// System API/SYS/API/bds_sys_do
///This function set the digital system output to the given state.
///
///=======
/// Remarks:
///=======
///    + The function is just used for the reactivation of the shunt after the elapsed recovery time and therefore a switch off is not necessary. 
///    + The |GVL_sys| is given for usage of defines.
///    + Import the bds_rts_ec.xml to use the enums. (Refer example below).
///
///----------
/// FFI:
///----------
///This API can be used in trusted partitions only. See Freedom from Interference (FFI) concept for more details.
///
///==================================================================		  			===================================================================================================
///Return value    								  									Description
///==================================================================		  			===================================================================================================
///16#00																				No error.
///16#01																				A parameter is invalid.
///16#02																				Function call was erroneous.
///16#03																				Shunt activation is not enabled.
///16#04																				Recovery time is not elapsed.
///
///==================================================================		   			===================================================================================================
///
///=======
///Code Example:
///=======
///============================================================================
///
///PROGRAM PLC_PRG
///
///VAR
///
///	status_u8: UISNT := 16#00; 
/// 
///	Init_flag_u8:USINT:=0;
///
///END_VAR
///
///  
///IF(Init_flag_u8=0) THEN (*To make api call once in application*)
///
///	(* reactivate the shunt after detection of a short circuit to battery *)
///	
///	status_u8 := bds_sys_do(bds_sys_do_signal_te.SHUNT1_EN, STD_ACTIVE);
///	
///	Init_flag_u8:=1;
///  
///END_IF
///
///============================================================================
{attribute 'external_name' := 'cmp_rts_bds_sys_do'}
FUNCTION bds_sys_do : USINT
VAR_INPUT
	///The assigned signal name.
	signal_e: UINT;
	///States of the sensor supply.
	///
	///    + STD_OFF - Disable the digital output,
	///    + STD_ON   - Enable the digital output.
	state_u8: USINT;
END_VAR

END_FUNCTION

// I/O API/IN legacy/API/bds_in_aid
///Get the analog voltage of the input as state.
///
///=======
/// Remarks:
///=======
///    + The evaluation of the state (and also the diagnosis OR (out of range)) is only possible with the configuration of the state thresholds. ( see |bds_in_aid_cfg|).
///
///----------
/// FFI:
///----------
///This API can be used in trusted partitions only. See Freedom from Interference (FFI) concept for more details.
///
///	
///==================================================================		  			===================================================================================================
///Return value    								  									Description
///==================================================================		  			===================================================================================================
///0																					No error
///1																					Invalid parameter
///2																					Function call was erroneous
///3																					Thresholds are not configured
///
///==================================================================		   			===================================================================================================
///
///=======
///Code Example:
///=======
///============================================================================
///
///PROGRAM appl_10ms_task
///  VAR
///  
///    stK59_u8: USINT := 16#00;
///  END_VAR
///
///  (* get the state of input K59 *)
///  
///  bds_in_aid(bds_in_aiv_signal_te.K59, ADR(stK59_u8));
///END
///
///============================================================================
{attribute 'external_name' := 'cmp_rts_bds_in_aid'}
FUNCTION bds_in_aid : USINT
VAR_INPUT
	///The signal name that is assigned to the respective pin configured as voltage input
	signal_e: UINT;
	///Storage address of the state.
	///	
	///States:
	///    + 0 : OFF
	///    + 1 : ON
	state_pu8: POINTER TO USINT;
END_VAR

END_FUNCTION

// I/O API/IN legacy/API/bds_in_aid_cfg
///Configure the state thresholds voltages of the input.
///
///=======
/// Remarks:
///=======
///    + The evaluation of the state and also the diagnosis of out of range (OR) is only possible with the configuration of the state thresholds (see also Configure a digital input.)
///	    + With a diagnosis threshold range of 150 to 4850mV or 150 to 19850mV or 150 to 39850mV, the corresponding state threshold range for the configurable inputs are defined from 300 to 4700mV or 300 to 19700mV or 300 to 39700mV depending upon the configuration.
///	    + With a diagnosis threshold range of 150 to 29850mV the state threshold range for the fixed inputs is defined from 300 to 29700mV. 
///    + For more information see |bds_in_aiv_getStatus|. 
///    + The AID_cfg  function is not recommended for the discrete inputs that have pull-up to battery (14K7) and pull-down (80K). 
///    + For discrete inputs, the thresholds depend on the battery voltage. It is recommended to do the evaluation of the states in ASW by reading the current battery voltage for a particular input and to calculate the appropriate thresholds for that battery voltage.
///
///----------
/// FFI:
///----------
///This API can be used in trusted partitions only. See Freedom from Interference (FFI) concept for more details.
///
///	
///==================================================================		  			===================================================================================================
///Return value    								  									Description
///==================================================================		  			===================================================================================================
///0																					No error
///1																					Invalid parameter
///
///==================================================================		   			===================================================================================================
///
///=======
///Code Example:
///=======
///============================================================================
///
///PROGRAM appl_10ms_task
///  VAR
///  
///  END_VAR
///
/// (* configure the state thresholds of input K59 *)
///
///  bds_in_aid_cfg(bds_in_aiv_signal_te.K59, 3000, 2000);
///END
///
///============================================================================
{attribute 'external_name' := 'cmp_rts_bds_in_aid_cfg'}
FUNCTION bds_in_aid_cfg : USINT
VAR_INPUT
	///The signal name that is assigned to the respective pin configured as voltage input
	signal_e: UINT;
	///Upper state threshold [mV].
	///
	///Range:
	///
	///Configurable inputs:
	///300 to 4700 / 300 to 19700 /300 to 39700
	///
	///Fixed inputs:
	///300 to 29700 
	///
	///Note:
	///upperThreshold_u16 > lowerThreshold_u16
	upperThreshold_u16: UINT;
	///Lower diagnosis threshold [mV].
	///
	///Range:
	///
	///Configurable inputs:
	///300 to 4700 / 300 to 19700 / 300 to 39700
	///
	///Fixed inputs:
	///300 to 29700
	///
	///Note:
	///lowerThreshold_u16 < upperThreshold_u16
	lowerThreshold_u16: UINT;
END_VAR

END_FUNCTION

// I/O API/IN legacy/API/bds_in_aiv
///Provides the analog voltage of the input.
///
///=======
/// Remarks:
///=======
///The voltage range of the inputs depends on the input type and the input configuration using eC (easyConfig). (see also |bds_in_aiv_cfg| and |bds_in_aid_cfg|).
///	   + Based on the configuration, the measurement range of the input  can  be  0 to 5000mV or 0 to 20000mV or 0 to 40000mV 
///	   + The measurement range of the routed input via the input device is 0 to 5000mV, see also Analog voltage aquisition.
///	   + The measurement range of the discrete inputs is 0 to 33000mV or 0 to 5000 mV
///
///
///----------
/// FFI:
///----------
///This API can be used in trusted partitions only. See Freedom from Interference (FFI) concept for more details.
///
///==================================================================		  			===================================================================================================
///Return value    								  									Description
///==================================================================		  			===================================================================================================
///0																					No error
///1																					Invalid parameter
///
///==================================================================		   			===================================================================================================
///
///
///=======
///Code Example:
///=======
///============================================================================
///
///PROGRAM appl_10ms_task
///  VAR
///  
///    mV_K59_u16: UINT := 16#00;
///  END_VAR
///
/// (* get the voltage of input K59 *)
///
///  bds_in_aiv(bds_in_aiv_signal_te.K59, ADR(mV_K59_u16));
///END
///
///============================================================================
{attribute 'external_name' := 'cmp_rts_bds_in_aiv'}
FUNCTION bds_in_aiv : USINT
VAR_INPUT
	///The signal name that is assigned to the respective pin configured as voltage input
	signal_e: UINT;
	///Storage address of the value.
	///
	///Range:
	///0 to 40000  [mV]
	value_pu16: POINTER TO UINT;
END_VAR

END_FUNCTION

// I/O API/IN legacy/API/bds_in_aiv_cfg
///Configures the diagnosis thresholds voltages of the input.
///
///=======
/// Remarks:
///=======
///   + The diagnosis is only possible after the configuration of the diagnosis thresholds. 
///	   + Depending on the configuration, the diagnosis threshold range for the configurable inputs can be from 150 to 4850 or 150 to 19850 or 150 to 39850mV.
///	   + The diagnosis threshold range for the fixed inputs ranges is from 150 to 29850mV or 150 to 4850 mV.
///   + For more information see |bds_in_aiv_getStatus|.
///   + This function should be called only once in the application.
///	
///
///----------
/// FFI:
///----------
///This API can be used in trusted partitions only. See Freedom from Interference (FFI) concept for more details.
///
///==================================================================		  			===================================================================================================
///Return value    								  									Description
///==================================================================		  			===================================================================================================
///0																					No error
///1																					Invalid parameter
///2																					Function call was erroneous.
///
///==================================================================		   			===================================================================================================
///
///=======
///Code Example:
///=======
///============================================================================
///
///PROGRAM PLC_PRG
///
///  VAR
///  
///	Init_flag_u8:USINT:=0;
/// 
///  END_VAR
///
///IF(Init_flag_u8=0) THEN (*To make api call once in application*)
///
///	(* configure diagnosis thresholds of input K59 *)
///	
///	bds_in_aiv_cfg(bds_in_aiv_signal_te.K59, 4850, 150);
///	
///	Init_flag_u8:=1;
///  
///END_IF
///
///============================================================================
{attribute 'external_name' := 'cmp_rts_bds_in_aiv_cfg'}
FUNCTION bds_in_aiv_cfg : USINT
VAR_INPUT
	///The signal name that is assigned to the respective pin configured as voltage input.
	signal_e: UINT;
	///Higher diagnosis threshold in [mV].
	///
	///Range:
	///
	///Configurable inputs:
	///150 to 4850 / 150 to 19850 / 150 to 39850
	///
	///Fixed inputs:
	///150 to 29850
	///
	///Note:
	///upperThreshold_u16 > lowerThreshold_u16
	upperThreshold_u16: UINT;
	///Lower diagnosis threshold in [mV].
	///
	///Range:
	///
	///Configurable inputs:
	///150 to 4850 / 150 to 19850 / 150 to 39850
	///
	///Fixed inputs:
	///150 to 29850
	///
	///Note:
	///lowerThreshold_u16 < upperThreshold_u16
	lowerThreshold_u16: UINT;
END_VAR

END_FUNCTION

// I/O API/IN legacy/API/bds_in_phase
///Provides the signal and the phase information of a channel (consist of a primary and a secondary frequency signal).
///
///=======
/// Remarks:
///=======
///   + The phase measurement for a phase channel can be configured through easyConfig and is automatically enabled during the start up of the ECU.
///   + All frequency inputs can be grouped to predefined input pairs.
///   + For information about the signal acquisition see Frequency aquisition.
///   + Following signal information is available: 
///	   + Frequency information of the primary signal [dHz].
///	   + Rotation direction information (0 = counter clockwise, 1 = clockwise).
///	   + The level of the secondary signal at rising edge of primary signal decides the rotation direction (signal low = 0 / signal high = 1).
///
///
///----------
/// FFI:
///----------
///This API can be used in trusted partitions only. See Freedom from Interference (FFI) concept for more details.
///
///
///==================================================================		  			===================================================================================================
///Return value    								  									Description
///==================================================================		  			===================================================================================================
///0																					No error
///1																					Invalid parameter
///2																					Function call was erroneous
///
///==================================================================		   			===================================================================================================
///
///
///=======
///Code Example:
///=======
///============================================================================
///
///PROGRAM appl_10ms_task
///
///   VAR
///   
///     phase_s: bds_in_phase_ts;
///	 
///     freq_u32: UDINT := 16#00;
///	 
///     dir_u8: USINT := 16#00;
///	 
///   END_VAR
///
///	(* phase measurement was activated within OsIniProc *)
///
///	bds_in_phase(bds_in_phase_signal_te.K54_VI_K37_VI, ADR(phase_s));
///
///	freq_u32 := phase_s.frequency_u32;
///
///	dir_u8   := phase_s.direction_u8;
///END
///
///============================================================================
{attribute 'external_name' := 'cmp_rts_bds_in_phase'}
FUNCTION bds_in_phase : USINT
VAR_INPUT
	///The signal name that is assigned to the respective pin configured as phase input
	signal_e: UINT;
	///Pointer to a structure |bds_in_phase_ts| with the phase information
	phase_ps: POINTER TO bds_in_phase_ts;
END_VAR

END_FUNCTION

// System API/DSM/API/bds_dsm_delErrorsJ1939
///This function is used to reset the status of all DFCs specified by the state and configured for J1939 only as well as to delete the related DFES entry if it exists.
///
///=======
/// Remarks:
///=======
///    + The |GVL_dsm| is given for usage of defines.
///	+ Suspect Parameter Number (SPN), Failure Mode Identifier (FMI) and Lamp States can be configured in easyConfig.
///
///----------
/// FFI:
///----------
///This API can be used in trusted partitions only. See Freedom from Interference (FFI) concept for more details.
///
///==================================================================		  			===================================================================================================
///Return value    								  									Description
///==================================================================		  			===================================================================================================
///16#0000: BDS_DSM_NO_ERROR_DU16														Update Number of Error is Successful .
///16#0004: BDS_DSM_INVALID_PTR_DU16													Invalid Pointer.
///16#0005: BDS_DSM_STATE_ERROR_DU16													Invalid State.
///
///==================================================================		   			===================================================================================================
///
///
///=======
///Code Example:
///=======
///============================================================================
///
///PROGRAM BDS_DSM_DEL_ERRORS__J1939_TEST
///
///VAR
///
///	status_u16: UINT;
///
///END_VAR
///
///dfc_s.id := dfc_ts.DFCid;
///
///(*Get the number of error*)
///
///status_u16 := bds_dsm_delErrorsJ1939(PREVIOUSLY_ACTIVE_ERRORS);
///
///if status_u16 = BDS_DSM_NO_ERROR_DU16 THEN
///
///	(*Error has been deleted successfully*)
///
///END_IF
///
///
///============================================================================
///
{attribute 'external_name' := 'cmp_rts_bds_dsm_delErrorsJ1939'}
FUNCTION bds_dsm_delErrorsJ1939 : UINT
VAR_INPUT
	///The kind of error status can be specified in detail by means of this mask.
	///	+ ACTIVE_ERRORS(0)                      - Fault is Active.
	///	+ PREVIOUSLY_ACTIVE_ERRORS(1) - Fault was Previously Active.
	state_e: bds_dsm_state_te;
END_VAR

END_FUNCTION

// System API/DSM/API/bds_dsm_delError_DTC
///This function resets the status of specific DFC as well as deletes the related DFES entry if it exists through DTC. 
///
///=======
/// Remarks:
///=======
///    + The |GVL_dsm| is given for usage of defines.
///
///----------
/// FFI:
///----------
///This API can be used in trusted partitions only. See Freedom from Interference (FFI) concept for more details.
///
///==================================================================		  			===================================================================================================
///Return value    								  									Description
///==================================================================		  			===================================================================================================
///16#0000: BDS_DSM_NO_ERROR_DU16														Both DFES entry and DFC status bit are cleared in DFC status memory.
///16#000B: BDS_DSM_NO_DTC_AVAILABLE_DU16												Invalid DTC.
///
///==================================================================		   			===================================================================================================
///
///
///=======
///Code Example:
///=======
///============================================================================
///
///PROGRAM BDS_DSM_DEL_ERROR_DTC_TEST
///
///VAR
///
///	status_u16: UINT;
///
///	dfc_s: bds_dsm_dfc_ts;	
///
///	dfc_ts : DFC_bds_NoDebFault1;
///
///END_VAR
///
///dfc_s.id := dfc_ts.DFCid;
///
///(*Deletes the Error status from DFC and related DFES entry*)
///
///status_u16 := bds_dsm_delError_DTC(dfc_ts.DTC); 
///
///if status_u16 = BDS_DSM_NO_ERROR_DU16 THEN
///
///	(*Error has been deleted successfully*)
///
///END_IF
///
///
///============================================================================
///
{attribute 'external_name' := 'cmp_rts_bds_dsm_delError_DTC'}
FUNCTION bds_dsm_delError_DTC : UINT
VAR_INPUT
	///DTC value : It is configured using easyConfig tool.
	dtc_u16: UINT;
END_VAR

END_FUNCTION

// I/O API/OUT_LEGACY/bds_out_poc_cfgPI
///Sets the gain values for Kp and Ki of a proportional output with current control.
///
///=======
/// Remarks:
///=======
///   + The range of Kp is defined as 0 to 2000 and for Ki as 0 to 500.
///   + The default values after reset of the ECU are Kp = 100 and Ki = 25.
///   + For more information see |bds_out_po_getStatus|.
///   + This function should be called only once in the application.
///
///----------
/// FFI:
///----------
///This API can be used in trusted partitions . For untrusted partitions use |bds_out_poc_cfgPI_ffi|. See Freedom from Interference (FFI) concept for more details.
///   
///==================================================================		  			===================================================================================================
///Return value    								  									Description
///==================================================================		  			===================================================================================================
///0																					No error.
///1																					A parameter is invalid.
///
///==================================================================		   			===================================================================================================
///
///=======
///Code Example:
///=======
///============================================================================
///
///PROGRAM PLC_PRG
///
///VAR
///
///	Init_flag_u8:USINT:=0;
///
///END_VAR
///  
///IF(Init_flag_u8=0) THEN (*To make api call once in application*)
///			
///	(* configure the gain values for output K73 *)
///	
///	bds_out_poc_cfgPI(bds_out_po_signal_te.K73, 200, 100);
///  
///	Init_flag_u8:=1;
///  
///END_IF
///
///============================================================================
{attribute 'external_name' := 'cmp_rts_bds_out_poc_cfgPI'}
FUNCTION bds_out_poc_cfgPI : USINT
VAR_INPUT
	///The connector assigned signal name of the output.
	signal_e: UINT;
	///Kp value.
	///
	///   + Range:0 to 2000
	///
	///   + Default : 100
	kp_u16: UINT;
	///Ki value. 
	///
	///   + Range:0 to 500
	///
	///   + Default : 25
	ki_u16: UINT;
END_VAR

END_FUNCTION

// I/O API/OUT/FFI_API/bds_out_poc_cfgPI_ffi
{attribute 'external_name' := 'cmp_rts_bds_out_poc_cfgPI_ffi'}
FUNCTION bds_out_poc_cfgPI_ffi : USINT
VAR_INPUT
	///The connector assigned signal name of the output.
	signal_e: UINT;
	///Kp value.
	///
	///   + Range:0 to 2000
	///
	///   + Default : 100
	kp_u16: UINT;
	///Ki value. 
	///
	///   + Range:0 to 500
	///
	///   + Default : 25
	ki_u16: UINT;
END_VAR

END_FUNCTION

// I/O API/IN legacy/API/bds_in_fi_cfg
///Configures the sensor type for a frequency input.
///
///=======
/// Remarks:
///=======
///   + The DSM frequency inputs support active sensors as well as DSM sensors and must therefore be configured according to the sensor type.
///   + For more information about the sensor types see |bds_in_fi|.
///   + For more  detailed information see |bds_in_fi_getStatus|.
///   + This function should be called only once in the application.
///
///----------
/// FFI:
///----------
///This API can be used in trusted partitions only. See Freedom from Interference (FFI) concept for more details.
///
///==================================================================		  			===================================================================================================
///Return value    								  									Description
///==================================================================		  			===================================================================================================
///0																					No error
///1																					Invalid parameter
///
///==================================================================		   			===================================================================================================
///
///
///=======
///Code Example:
///=======
///============================================================================
///
///PROGRAM PLC_PRG
///
///  VAR
///  
///	Init_flag_u8:USINT:=0;
/// 
///  END_VAR
///  
///IF(Init_flag_u8=0) THEN (*To make api call once in application*)
///
///	(* DSM sensor is used for input K37_VI *)
///	
///	bds_in_fi_cfg(bds_in_fi_signal_te.K37_VI, STD_ON);
///	
///	(* active sensor is used for input K61_VI *)
///	
///	bds_in_fi_cfg(bds_in_fi_signal_te.K61_VI, STD_OFF);
///  
///	Init_flag_u8:=1;
///  
///END_IF
///
///============================================================================
{attribute 'external_name' := 'cmp_rts_bds_in_fi_cfg'}
FUNCTION bds_in_fi_cfg : USINT
VAR_INPUT
	///The signal name that is assigned to the respective pin configured as frequency input
	signal_e: UINT;
	///Configuration of the sensor type.
	///   + STD_OFF - Active sensor
	///   + STD_ON   - DSM sensor
	dsmSensor_u8: USINT;
END_VAR

END_FUNCTION

// I/O API/IN legacy/API/bds_in_fi
///Provides the frequency of the input.
///
///=======
/// Remarks:
///=======
///   + The measurement range of the frequency [dHz] is defined from 1 to 20 kHz. 
///   + To get the status of the input use |bds_in_fi_getStatus|.
///   + The DSM frequency inputs support active sensors as well as DSM sensors (see RE 95132). Therefore the DSM frequency inputs must be configured for  a particular sensor type using |bds_in_fi_cfg|. If a DSM sensor is used in an application, the shunt should be activated using easyConfig. A logical OR operation is performed on the  additional direction and status info of a DSM sensor and the frequency.
///   + In order to mask the info, it is mandatory to use the macros  BODAS API library, bds_rts_ec.xml (see example below).
///
///   + The format of frequency data is shown below (see the example below):
///   
///	   + 16#FFFFFFFF where, 
///			+ First two 'F'->status DSM sensor
///			+ Third letter 'F' -> direction DSM sensor
///			+ Last five letter 'F'->frequency
///   + If the situations where a DSM sensor is used, the shunt must be protected against the current values that exceeds 24000µA. Further, after the deactivation of shunt, a recovery time of 2s is required. 
///   + After the recovery time elapses, the shunt configuration can be enabled again using |bds_sys_do|.
///   + For more info about the shunt protection see |bds_in_fi_getStatus|.
///
///
///----------
/// FFI:
///----------
///This API can be used in trusted partitions only. See Freedom from Interference (FFI) concept for more details.
///
///==================================================================		  			===================================================================================================
///Return value    								  									Description
///==================================================================		  			===================================================================================================
///0																					No error
///1																					Invalid parameter
///2																					Function call was erroneous.
///
///==================================================================		   			===================================================================================================
///
///
///=======
///Code Example:
///=======
///============================================================================
///
///PROGRAM PLC_PRG
///
///  VAR
///  
///	Init_flag_u8:USINT:=0;
/// 
///  END_VAR
///  
///IF(Init_flag_u8=0) THEN (*To make api call once in application*)
///
///	(* Precondition for the use of a DSM sensor 
///	 * - shunt at the input shall be activated (configured with eC) and
///	 * - configured for a DSM sensor 
///	 * at start up. *)
///	
///	bds_in_fi_cfg(bds_in_fi_signal_te.K55_VI, STD_ACTIVE);
///  
///	Init_flag_u8:=1;
///  
///END_IF
///
///PROGRAM appl_10ms_task
///  VAR
///		fK53_u32: UDINT := 16#00;
///		fDSM_K55_u32: UDINT := 16#00;
///		fDSM_u32: UDINT := 16#00;
///		stDSM_u32: UDINT := 16#00;
///		dirDSM_u32: UDINT := 16#00;
///  END_VAR
///
///(* w/o preconditions *)
///   bds_in_fi(bds_in_fi_signal_te.K53, ADR(fK53_u32));
///
///(* preconditions for DSM sensor set in OsIniProc *)
///
///   bds_in_fi(bds_in_fi_signal_te.K55_VI, ADR(fDSM_K55_u32));
///
///(* get frequency, status and direction of DSM sensor *)
///
///  fDSM_u32   := fDSM_K55_u32 AND maskFrequency_DU32;
///  
///  stDSM_u32  := SHR((fDSM_K55_u32 AND maskStatus_DU32), numShiftStatus_DU32);
///  
///  dirDSM_u32 := SHR((fDSM_K55_u32 AND maskDirection_DU32), numShiftDirection_DU32);
///  
///END
///
///============================================================================
{attribute 'external_name' := 'cmp_rts_bds_in_fi'}
FUNCTION bds_in_fi : USINT
VAR_INPUT
	///The signal name that is assigned to the respective pin configured as frequency input
	signal_e: UINT;
	///Storage address of the value.
	///
	///Frequency [Nibbles 0...4]:
	///0..200000 [0,1Hz]
	///
	///Additional information if a DSM sensor is used.
	///
	///Direction [Nibble 5]:
	///   + 16#00 - standstill
	///   + 16#01 - left
	///   + 16#02 - right
	///   + 16#04 - unknown
	///
	///Status [Nibble 6...7]:
	///   + 16#00 - error free
	///   + 16#01 - air gap error 
	///   + 16#02 - mounting error
	///   + 16#04 - undefined signal length
	///   + 16#08 - period too long or measured period exceeds maximum period
	///   + 16#10 - no status signal available
	fi_pu32: POINTER TO UDINT;
END_VAR

END_FUNCTION

// I/O API/IN legacy/API/bds_in_fi_getStatus
///Provides the status of the input.
///
///=======
/// Remarks:
///=======
///   + For information about the signal acquisition see Frequency aquisition.
///   + The status data provides all relevant information about the frequency input (see the example below). 
///   + The structure member status_b16 holds the information regarding the configuration (see also |bds_in_fi_cfg|) and the shunt status of the DSM frequency input.
///   + A pulse counter of 15 bits is supported.
///
///----------
/// FFI:
///----------
///This API can be used in trusted partitions only. See Freedom from Interference (FFI) concept for more details.
///
///-----
/// INFO:
///----- 
///The special input circuit of the DSM frequency inputs also allows the input levels to be monitored additionally by configuring the corresponding diagnostic thresholds of the analog inputs.
///
///Example of an analog current input:
///
///In the example below K55_VI is used  for a DSM sensor. Due to the current interface (the current values are iHigh  = 14mA and iLow = 7mA) the analog current input can be used for an additional signal check. 
///If  current thresholds are configured  then it is possible to detect  short circuit to ground faults.
///A short circuit to battery leads to a deactivation of the shunt (shunt protection is faster than the diagnostic check.
///
///bds_in_aic_cfg(bds_in_fi_signal_te.K55_VI, 18000, 3000);
///bds_in_aic_getStatus(bds_in_fi_signal_te.K55_VI, ADR(stInK55_s));
///
///Also an analog voltage input can be used:
///
///bds_in_aiv_cfg(bds_in_fi_signal_te.K55, 3600, 600);
///bds_in_aiv_getStatus(bds_in_fi_signal_te.K55, ADR(stInK55_s));
///
///
///==================================================================		  			===================================================================================================
///Return value    								  									Description
///==================================================================		  			===================================================================================================
///0																					No error
///1																					Invalid parameter
///
///==================================================================		   			===================================================================================================
///
///
///
///=======
///Code Example:
///=======
///============================================================================
///
///PROGRAM PLC_PRG
///
///  VAR
///  
///	Init_flag_u8:USINT:=0;
/// 
///  END_VAR
///  
///IF(Init_flag_u8=0) THEN (*To make api call once in application*)
///
///	(* Precondition for the use of a DSM sensor
///	* - shunt at the input shall be activated (configured with eC) and
///	* - configured for a DSM sensor 
///	* at start up. *)
///	
///	bds_in_fi_cfg(bds_in_fi_signal_te.K55_VI, STD_ACTIVE);
///	
///	Init_flag_u8:=1;
///  
///END_IF
///
///PROGRAM appl_10ms_task
///   VAR
///   
///     stK53_s: bds_in_fi_ts;
///	 
///     fDSM_K55_u32: bds_in_fi_ts;
///	 
///   END_VAR
///
/// (* get the status of input K53 *)
/// 
///	bds_in_fi_getStatus(bds_in_fi_signal_te.K53, ADR(stK53_s));
///
/// (* get the status of input K55_VI *)
/// 
///	bds_in_fi_getStatus(bds_in_fi_signal_te.K55_VI, ADR(fDSM_K55_u32));
///	
///END
///
///============================================================================
{attribute 'external_name' := 'cmp_rts_bds_in_fi_getStatus'}
FUNCTION bds_in_fi_getStatus : USINT
VAR_INPUT
	///The signal name that is assigned to the respective pin configured as frequency input
	signal_e: UINT;
	///Storage address of the data.
	data_ps: POINTER TO bds_in_fi_ts;
END_VAR

END_FUNCTION

// I/O API/IN legacy/API/bds_in_phase_getStatus
///Provides information about the entities related to  phase measurement. For example frequency, direction, periods, time stamps, phase, pulse counter and the error status of a channel (consists of a primary and a secondary frequency signal).
///
///The bds_in_phase_getStatus API function get the data of the extended frequency acquisition.
///
///=======
/// Remarks:
///=======
///   + The phase measurement for a phase channels can be configured with eC and is automatically enabled during the start up of the ECU.
///   + For information about the signal acquisition see Frequency acquisition.
///   + If the application calls this function with an invalid channel parameter then the contents of the associated data structure will be 0.
///   + Following signal information is available: 
///	   + Frequency information                   
///	   + Direction of rotation (0 = counter clockwise, 1 = clockwise).
///	   + With respect to the error status of primary and secondary signal,  a failure in either of the signal is only detected if  both primary and secondary signals are available. 
///	   + Period [us] of the primary signal. 
///	   + Period [us] of the secondary signal. (The secondary signal is sometimes inconsistent)
///	   + Time stamp [us] of rising edge of the primary signal.
///	   + Time stamp [us] of rising edge of the secondary signal.
///	   + Phase shift [us] between the primary and the secondary signal (calculation is tiShift_u32 = tiSecSig_u32 - tiPrimSig_u32).
///	   + Pulse counter has  a resolution of +/- 2^23 .Pulses are counted with the rising edge with respect to the primary signal. 
///	   + The direction of counting also depends on the state of the secondary signal with respect to  the rising edge of the primary signal:  
///			   + 0 = increment
///			   + 1 = decrement 
///   + Signal state of the primary signal: 
///	   + state at function call time ("1" for high or "0" for low)
///	   + no update available (request with the same period)
///	   + period too long (timer overflow)
///	   + max-period exceeds given maximum length
///   + Signal state of the secondary signal:
///	   + state at function call time ("1" for high or "0" for low)
///	   + no update available (request with the same period)
///	   + period too long (timer overflow)
///	   + max-period exceeds given maximum length.
///   + The pulse counter can be reset with function |bds_in_phase_resetCounter|.
///   + Pointer to the start address of the Period array (size Max 20) for each signal is available for both the signals (primary and secondary). Further explanation of the extended frequency acquisition could be found under Frequency acquisition. 
///   + Pointer to the start address of Pulse array (size Max 20) is only available for the primary signal. Further explanation of the extended frequency acquisition could be found under Frequency acquisition. 
///   + As soon as the function is called, the data could be used within a loop, which will go over the 20 addresses in order to get all the contents of the array.
///   + Max-Period of the the primary signal must be configured with eC. The secondary signal will get the Max-Period value from the primary signal. 
///   + The Max-Period is set to 1 second (Default value on eC) and can be reduced to 1 millisecond.
///
///
///----------
/// FFI:
///----------
///This API can be used in trusted partitions only. See Freedom from Interference (FFI) concept for more details.
///
///==================================================================		  			===================================================================================================
///Return value    								  									Description
///==================================================================		  			===================================================================================================
///0																					No error
///1																					Invalid parameter
///2																					Function call was erroneous
///
///==================================================================		   			===================================================================================================
///
///
///
///=======
///Code Example:
///=======
///============================================================================
///
///PROGRAM appl_10ms_task
///   VAR
///   
///     stPhase_s: bds_in_stPhase_ts;
///	 
///     tiPeriodPrim_u32: UDINT := 16#00;
///	 
///     tiPeriodSec_u32: UDINT := 16#00;
///	 
///     tiShift_u32: UDINT := 16#00;
///	 
///   END_VAR
///
///  (* phase measurement is activated with the eC configuration *)
///  
///  bds_in_phase_getStatus(bds_in_phase_signal_te.K54_VI_K37_VI, ADR(stPhase_s));
///
///  (* get periods and phase position of signals *)
///  
///  tiPeriodPrim_u32 := stPhase_s.tiPeriodPrimSig_u32;
///  
///  tiPeriodSec_u32  := stPhase_s.tiPeriodSecSig_u32;
///  
///  tiShift_u32      := stPhase_s.tiShift_u32;
///END
///
///============================================================================
{attribute 'external_name' := 'cmp_rts_bds_in_phase_getStatus'}
FUNCTION bds_in_phase_getStatus : USINT
VAR_INPUT
	///The signal name that is assigned to the respective pin configured as phase input
	signal_e: UINT;
	///Pointer to the data structure |bds_in_stPhase_ts|
	stPhase_ps: POINTER TO bds_in_stPhase_ts;
END_VAR

END_FUNCTION

// I/O API/IN legacy/API/bds_in_phase_resetCounter
///Resets the directional pulse counter of a phase channel. It consists of a primary and a secondary frequency channel.
///
///=======
/// Remarks:
///=======
///   + The phase measurement for a phase channel can be configured using eC and is automatically enabled during the start up of the ECU.
///   + More information about the directional pulse counter can be found in the description at |bds_in_phase_getStatus|.
///
///
///----------
/// FFI:
///----------
///This API can be used in trusted partitions only. See Freedom from Interference (FFI) concept for more details.
///
///==================================================================		  			===================================================================================================
///Return value    								  									Description
///==================================================================		  			===================================================================================================
///0																					No error
///1																					Invalid parameter
///2																					Function call was erroneous
///
///==================================================================		   			===================================================================================================
///
///
///=======
///Code Example:
///=======
///============================================================================
///
///
///	VAR_GLOBAL
///	
///	   (* global variable *)
///	   
///	   pulseCounter_s32: DINT := 16#00;
///	   
///	END_VAR
///
///(* Read the position of a steering wheel using the pulse counter. Pulse counter is synchronized at null position *)
///
///PROGRAM appl_10ms_task
///   VAR
///   
///     stPhase_s: bds_in_stPhase_ts;
///	 
///     stK42_u8: USINT := 16#00;
///	 
///   END_VAR
///
/// (* check for null position of the steering wheel via digital input K42 *)
/// 
/// 	bds_in_di(bds_in_di_signal_te.K42, ADR(stK42_u8));
///
/// 	IF (1 == stK42_u8) THEN
///	
///   		(* reset the pulse counter if null position of steering wheel is detected *)
///		
///   		bds_in_phase_resetCounter(bds_in_phase_signal_te.K54_VI_K37_VI);
///		
/// 	END_IF
///
///   (* get data from phase measurement *)
///   
///   bds_in_phase_getStatus(bds_in_phase_signal_te.K54_VI_K37_VI, ADR(stPhase_s));
///
///   (* read pulse counter value *)
///   
///   pulseCounter_s32 := stPhase_s.couPulse_s32;
///END
///
///============================================================================
{attribute 'external_name' := 'cmp_rts_bds_in_phase_resetCounter'}
FUNCTION bds_in_phase_resetCounter : USINT
VAR_INPUT
	///The signal name that is assigned to the respective pin configured as phase input
	signal_e: UINT;
END_VAR

END_FUNCTION

// I/O API/IN legacy/API/bds_in_di
///Provides the digital state of the input.
///
///=======
/// Remarks:
///=======
///   + Thresholds for bds_in_di are not configured in the API. But, there are three pairs of theresholds that can be selected in configuration tool easyConfig.
///
///----------
/// FFI:
///----------
///This API can be used in trusted partitions only. See Freedom from Interference (FFI) concept for more details.
///
///==================================================================		  			===================================================================================================
///Return value    								  									Description
///==================================================================		  			===================================================================================================
///0																					No error
///1																					Invalid parameter
///2																					Function call was erroneous.
///
///==================================================================		   			===================================================================================================
///
///=======
///Code Example:
///=======
///============================================================================
///
///PROGRAM appl_10ms_task
///  VAR
///  
///    stK42_u8: USINT := 16#00;
///	
///  END_VAR
///
///  (* get the state of input K42 *)
///  
///  bds_in_di(bds_in_di_signal_te.K42, ADR(stK42_u8));
///  
///END
///
///============================================================================
{attribute 'external_name' := 'cmp_rts_bds_in_di'}
FUNCTION bds_in_di : USINT
VAR_INPUT
	///The signal name that is assigned to the respective pin configured as digital input
	signal_e: UINT;
	///Storage address of the state.
	///
	///States:
	///0 : OFF
	///1 : ON
	state_pu8: POINTER TO USINT;
END_VAR

END_FUNCTION

// I/O API/OUT_LEGACY/bds_out_po_cfgPwrLs
///Configures a proportional high side output as power supply for the low side outputs.
///
///=======
/// Remarks:
///=======
///   + The output is also switched on with the configuration.
///   + If the output is switched off and switched on again with |bds_out_pod| the open load faults of the connected low sides must be reset with |bds_out_po_resetError| respective |bds_out_do_resetError|.
///   + A high side output must be used for the power supply of the low sides because a direct supply of the low side outputs is not permitted.
///   + If the low side K51 shall be used as a proportional output, a power supply by a high side output is necessary.
///   + This function should be called only once in the application.
///
///----------
/// FFI:
///----------
///This API can be used in trusted partitions . For untrusted partitions use |bds_out_po_cfgPwrLs_ffi|. See Freedom from Interference (FFI) concept for more details.
///   
///------
/// Info:
///------
///
///With the configuration the open load detection is suppressed for the high side output. Therefore the output shall be configured during the start up of the RC, otherwise a fault may be detected depending on the time of configuration.
///
///==================================================================		  			===================================================================================================
///Return value    								  									Description
///==================================================================		  			===================================================================================================
///0																					No error.
///1																					A parameter is invalid.
///2																					Function call was erroneous.
///3																					Already configured as POC.
///4																					Output is disabled.
///5																					Output is locked
///6																					Output is already configured
///
///==================================================================		   			===================================================================================================
///
///=======
///Code Example:
///=======
///============================================================================
///
///PROGRAM PLC_PRG
///
///VAR
///
///	Init_flag_u8:USINT:=0;
///
///END_VAR
///  
///IF(Init_flag_u8=0) THEN (*To make api call once in application*)
///				
///	(* configure  proportional output as power supply for the low sides *)
///	
///	bds_out_po_cfgPwrLs(bds_out_po_signal_te.K09);
///  
///	Init_flag_u8:=1;
///  
///END_IF
///
///
///PROGRAM appl_10ms_task
///
///VAR
///
///END_VAR
///
///
///(* set duty cycle at high power output K51 *)
///
///bds_out_po(bds_out_po_signal_te.K51, 250);
///
///
///
///(* set duty cycle and state at low power outputs K80 and K84 *)
///
///bds_out_po(bds_out_po_signal_te.K80, 500);
///
///bds_out_do(bds_out_po_signal_te.K84, STD_ACTIVE);
///
///============================================================================
{attribute 'external_name' := 'cmp_rts_bds_out_po_cfgPwrLs'}
FUNCTION bds_out_po_cfgPwrLs : USINT
VAR_INPUT
	///The connector assigned signal name of the high side output
	signal_e: UINT;
END_VAR

END_FUNCTION

// I/O API/OUT_LEGACY/bds_out_pod
///Sets the proportional output to a state.
///
///=======
/// Remarks:
///=======
///
///   + The proportional output is controlled digitally .
///   + For more information see |bds_out_po_getStatus| and |bds_out_po_resetError|.
///
///
///----------
/// FFI:
///----------
///This API can be used in trusted partitions . For untrusted partitions use |bds_out_pod_ffi|. See Freedom from Interference (FFI) concept for more details.
///
///==================================================================		  			===================================================================================================
///Return value    								  									Description
///==================================================================		  			===================================================================================================
///0																					No error.
///1																					A parameter is invalid.
///2																					Function call was erroneous.
///3																					Already configured as POC.
///4																					Output is disabled.
///5																					Output is locked
///6																					Already configured as SAFOUT channel
///
///==================================================================		   			===================================================================================================
///
///=======
///Code Example:
///=======
///============================================================================
///
///PROGRAM appl_10ms_task
///
///VAR
///
///END_VAR
///
///(* activate proportional output with digital state *)
///
///bds_out_pod(bds_out_po_signal_te.K73, STD_ACTIVE);
///
///============================================================================
{attribute 'external_name' := 'cmp_rts_bds_out_pod'}
FUNCTION bds_out_pod : USINT
VAR_INPUT
	///The connector assigned signal name of the output.
	signal_e: UINT;
	///State of the output.
	///   + STD_IDLE
	///   + STD_ACTIVE
	state_u8: USINT;
END_VAR

END_FUNCTION

// I/O API/OUT/FFI_API/bds_out_pod_ffi
{attribute 'external_name' := 'cmp_rts_bds_out_pod_ffi'}
FUNCTION bds_out_pod_ffi : USINT
VAR_INPUT
	///The connector assigned signal name of the output.
	signal_e: UINT;
	///State of the output.
	///   + STD_IDLE
	///   + STD_ACTIVE
	state_u8: USINT;
END_VAR

END_FUNCTION

// I/O API/OUT/FFI_API/bds_out_po_cfgPwrLs_ffi
{attribute 'external_name' := 'cmp_rts_bds_out_po_cfgPwrLs_ffi'}
FUNCTION bds_out_po_cfgPwrLs_ffi : USINT
VAR_INPUT
	///The connector assigned signal name of the high side output
	signal_e: UINT;
END_VAR

END_FUNCTION

// I/O API/SAFOUT/API/bds_safout_resetError
///Resets errors of a channel.
///
///=======
/// Remarks:
///=======
///   + The fault status of all outputs is reset as well as the DFC of the channel.
///   + For more information see Linked outputs.
///
///----------
/// FFI:
///----------
///This API can be used in trusted partitions only. See Freedom from Interference (FFI) concept for more details.
///
///-----
/// Info:
///-----
///
///After a fault the channel is switched off and locked. A call to |bds_safout_resetError| is the precondition for unlocking  the channel. Also see  |bds_safout_unlock|. Resetting the errors takes some time, therefore a delay is necessary for calling the unlock function.
///
///==================================================================		  			===================================================================================================
///Return value    								  									Description
///==================================================================		  			===================================================================================================
///0																					No error.
///1																					A parameter is invalid.
///
///==================================================================		   			===================================================================================================
///
///=======
///Code Example:
///=======
///============================================================================
///
///VAR_GLOBAL CONSTANT
///
///   (* safout channel name *)
///
///   PHDLS_CHNL1: UINT := (PHDLS OR CHNL1);
///
///   DHDLM_CHNL2: UINT := (DHDLM OR CHNL2);
///
///   PHMDL_CHNL3: UINT := (PHMDL OR CHNL3);
///
///END_VAR
///
/// 
///PROGRAM PLC_PRG
///
///VAR
///
///END_VAR
///
///
///
///(* configure for POC *)
///
///bds_out_po_cfg(bds_out_po_signal_te.K73, STD_ACTIVE);
///
///bds_out_po_cfg(bds_out_po_signal_te.K07, STD_ACTIVE);
///
///bds_out_po_cfg(bds_out_po_signal_te.K29, STD_ACTIVE);
///
///bds_out_po_cfg(bds_out_po_signal_te.K09, STD_ACTIVE);
///
///
///
///(* configure channels for SAFOUT *)
///
///bds_safout_cfg(PHDLS_CHNL1, bds_out_po_signal_te.K73, bds_out_po_signal_te.K51, bds_out_do_signal_te.K14, 0, 0);
///
///bds_safout_cfg(DHDLM_CHNL2, bds_out_po_signal_te.K08, bds_out_do_signal_te.K16, bds_out_do_signal_te.K15, bds_out_do_signal_te.K13, 0);
///
///bds_safout_cfg(PHMDL_CHNL3, bds_out_do_signal_te.K12, bds_out_po_signal_te.K07, bds_out_po_signal_te.K29, bds_out_po_signal_te.K09, 0);
///
///
///
///PROGRAM appl_10ms_task
///
///VAR
///
///END_VAR
///
///
///(* reset channels *)
///
///bds_safout_resetError(PHDLS_CHNL1);
///
///bds_safout_resetError(DHDLM_CHNL2);
///
///bds_safout_resetError(PHMDL_CHNL3);
///
///============================================================================
{attribute 'external_name' := 'cmp_rts_bds_safout_resetError'}
FUNCTION bds_safout_resetError : USINT
VAR_INPUT
	///The connector assigned signal name of the output.
	///
	///The channel name is composed of mode and channel number
	///
	///channel name = mode OR channel number
	///
	///and shall be defined from the application (see also example below):
	///
	///PHDLS_CHNL1: UINT := (PHDLS OR CHNL1)
	chnl_u16: UINT;
END_VAR

END_FUNCTION

// I/O API/SAFOUT/API/bds_safout_unlock
///Unlocks a locked channel.
///
///=======
/// Remarks:
///=======
///
///   + When cause of a fault has been corrected  then first reset the errors using |bds_safout_resetError|  and then unlock the safeout channel for further usage.  See also |bds_safout_ignoreError|.
///   + Resets frozen diagnostic value in |bds_safout_getStatus|.  
///
///
///----------
/// FFI:
///----------
///This API can be used in trusted partitions only. See Freedom from Interference (FFI) concept for more details.
///
///==================================================================		  			===================================================================================================
///Return value    								  									Description
///==================================================================		  			===================================================================================================
///0																					No error.
///1																					A parameter is invalid.
///2																					Errors are not reset.
///
///==================================================================		   			===================================================================================================
///
///=======
///Code Example:
///=======
///============================================================================
///
///VAR_GLOBAL CONSTANT
///
///   (* safout channel name *)
///
///   PHDLS_CHNL1: UINT := (PHDLS OR CHNL1);
///
///   DHDLM_CHNL2: UINT := (DHDLM OR CHNL2);
///
///   PHMDL_CHNL3: UINT := (PHMDL OR CHNL3);
///
///END_VAR
///
/// 
///
///PROGRAM PLC_PRG
///
///VAR
///
///END_VAR
///
///
///
///(* configure for POC *)
///
///bds_out_po_cfg(bds_out_po_signal_te.K73, STD_ACTIVE);
///
///bds_out_po_cfg(bds_out_po_signal_te.K07, STD_ACTIVE);
///
///bds_out_po_cfg(bds_out_po_signal_te.K29, STD_ACTIVE);
///
///bds_out_po_cfg(bds_out_po_signal_te.K09, STD_ACTIVE);
///
///
///
///(* configure channels for SAFOUT *)
///
///bds_safout_cfg(PHDLS_CHNL1, bds_out_po_signal_te.K73, bds_out_po_signal_te.K51, bds_out_do_signal_te.K14, 0, 0);
///
///bds_safout_cfg(DHDLM_CHNL2, bds_out_po_signal_te.K08, bds_out_do_signal_te.K16, bds_out_do_signal_te.K15, bds_out_do_signal_te.K13, 0);
///
///bds_safout_cfg(PHMDL_CHNL3, bds_out_do_signal_te.K12, bds_out_po_signal_te.K07, bds_out_po_signal_te.K29, bds_out_po_signal_te.K09, 0);
///
///
///PROGRAM appl_10ms_task
///
///VAR
///
///END_VAR
///
///
///
///(* reset channels *)
///
///bds_safout_unlock(PHDLS_CHNL1);
///
///bds_safout_unlock(DHDLM_CHNL2);
///
///bds_safout_unlock(PHMDL_CHNL3);
///
///
///============================================================================
{attribute 'external_name' := 'cmp_rts_bds_safout_unlock'}
FUNCTION bds_safout_unlock : USINT
VAR_INPUT
	///The connector assigned signal name of the output.
	///
	///The channel name is composed of mode and channel number
	///
	///channel name = mode OR channel number
	///
	///and shall be defined from the application (see also example below):
	///
	///PHDLS_CHNL1: UINT := (PHDLS OR CHNL1)
	chnl_u16: UINT;
END_VAR

END_FUNCTION

// I/O API/SAFOUT/API/bds_safout_ignoreError
///Ignores errors, that only affect the capability to shutdown a channel.
///
///=======
/// Remarks:
///=======
///   + This feature is valid only for PHMDL, PLMDH, DHDLM and DLDHM mode. 
///   + To increase availability, faults that only affect the capability to shutdown a channel can be ignored and the channel is released again. The configuration is not saved, therefore the fault is only ignored until the next reset of the ECU, or the ignoring is canceled by the application.
///   + This function also ignores the current deviation errors, i.e., safout channel is not locked but current deviation DFC is set, if error occurred. 
///
///----------
/// FFI:
///----------
///This API can be used in trusted partitions only. See Freedom from Interference (FFI) concept for more details.
///
///-----
/// Danger:
///-----
///
///The use of the function has an impact for the functional safety.
///
///==================================================================		  			===================================================================================================
///Return value    								  									Description
///==================================================================		  			===================================================================================================
///0																					No error.
///1																					A parameter is invalid.
///2																					wrong mode or channel
///3																					Feature is not supported of this mode
///
///==================================================================		   			===================================================================================================
///
///=======
///Code Example:
///=======
///============================================================================
///
///VAR_GLOBAL CONSTANT
///
///   (* safout channel name *)
///
///   PHDLS_CHNL1: UINT := (PHDLS OR CHNL1);
///
///   DHDLM_CHNL2: UINT := (DHDLM OR CHNL2);
///
///   PHMDL_CHNL3: UINT := (PHMDL OR CHNL3);
///   
///   PLDHS_CHNL4: UINT := (PLDHS OR CHNL4);
///
///   DLDHM_CHNL5: UINT := (DLDHM OR CHNL5);
///
///   PLMDH_CHNL6: UINT := (PLMDH OR CHNL6);
///
///END_VAR
///
/// 
///
///PROGRAM PLC_PRG
///
///VAR
///
///END_VAR
///
///
///
///(* configure for POC *)
///
///bds_out_po_cfg(bds_out_po_signal_te.K73, STD_ACTIVE);
///
///bds_out_po_cfg(bds_out_po_signal_te.K07, STD_ACTIVE);
///
///bds_out_po_cfg(bds_out_po_signal_te.K29, STD_ACTIVE);
///
///bds_out_po_cfg(bds_out_po_signal_te.K09, STD_ACTIVE);
///
///
///
///(* configure channels for SAFOUT *)
///
///bds_safout_cfg(PHDLS_CHNL1, bds_out_po_signal_te.K73, bds_out_po_signal_te.K51, bds_out_do_signal_te.K14, 0, 0);
///
///bds_safout_cfg(DHDLM_CHNL2, bds_out_po_signal_te.K08, bds_out_do_signal_te.K16, bds_out_do_signal_te.K15, bds_out_do_signal_te.K13, 0);
///
///bds_safout_cfg(PHMDL_CHNL3, bds_out_do_signal_te.K12, bds_out_po_signal_te.K07, bds_out_po_signal_te.K29, bds_out_po_signal_te.K09, 0);
///
///bds_safout_cfg(PLDHS_CHNL4, bds_out_po_signal_te.A19, bds_out_po_signal_te.A32, bds_out_do_signal_te.A47, 0, 0);
///
///bds_safout_cfg(DLDHM_CHNL5, bds_out_po_signal_te.A03, bds_out_do_signal_te.A33, bds_out_do_signal_te.A46, bds_out_do_signal_te.A48, 0);
///
///bds_safout_cfg(PLMDH_CHNL6, bds_out_do_signal_te.A31, bds_out_po_signal_te.A05, bds_out_po_signal_te.A20, 0, 0);
///
///
///PROGRAM appl_10ms_task
///
///VAR
///
///END_VAR
///
///
///
///(* ignore existing faults *)
///
///bds_safout_ignoreError(PHDLS_CHNL1, STD_ON);
///
///bds_safout_ignoreError(DHDLM_CHNL2, STD_ON);
///
///bds_safout_ignoreError(DLDHM_CHNL5, STD_ON);
///
///bds_safout_ignoreError(PLMDH_CHNL6, STD_ON);
///
///(* existing fault is no longer ignored, example to switch OFF ignore error feature*)
///
///bds_safout_ignoreError(PHDLS_CHNL1, STD_OFF);
///
///
///============================================================================
{attribute 'external_name' := 'cmp_rts_bds_safout_ignoreError'}
FUNCTION bds_safout_ignoreError : USINT
VAR_INPUT
	///The connector assigned signal name of the output.
	///
	///The channel name is composed of mode and channel number
	///
	///channel name = mode OR channel number
	///
	///and shall be defined from the application (see also example below):
	///
	///PHDLS_CHNL1: UINT := (PHDLS OR CHNL1)
	chnl_u16: UINT;
	///Select, if the error shall be ignored
	///
	///State: STD_OFF(16#00) or STD_ON(16#01) 
	state_u8: USINT;
END_VAR

END_FUNCTION

// I/O API/SAFOUT/API/bds_safout_cfg
///Configures a channel with the desired mode.
///
///=======
/// Remarks:
///=======
///   + A channel shall be configured with ECU specific modes.
///   + With the available resources of the RC27-18/40, up to 18 channels and the RC18-12/40 up to 12 channels can be configured.
///   + Parameters out1_u16 to out4_u16 shall be configured in an ascending order.
///   + For unused output parameters a "0" shall be used.
///   + Dependent from the desired mode, the proportional output(s) shall be configured as first as POC, see |bds_out_po_cfg|.
///   + For more information, see also |bds_safout_getStatus|.
///
///----------
/// FFI:
///----------
///This API can be used in trusted partitions only. See Freedom from Interference (FFI) concept for more details.
///
///==================================================================		  			===================================================================================================
///Return value    								  									Description
///==================================================================		  			===================================================================================================
///0																					No error.
///1																					A parameter is invalid.
///2																					outCo is already configured
///3																					out1 is already configured
///4																					out2 is already configured
///5																					out3 is already configured
///6																					out4 is already configured
///
///==================================================================		   			===================================================================================================
///
///=======
///Code Example:
///=======
///============================================================================
///
///VAR_GLOBAL CONSTANT
///
///   (* safout channel name *)
///
///   PHDLS_CHNL1: UINT := (PHDLS OR CHNL1);
///
///   DHDLM_CHNL2: UINT := (DHDLM OR CHNL2);
///
///   PHMDL_CHNL3: UINT := (PHMDL OR CHNL3);
///   
///   PLDHS_CHNL4: UINT := (PLDHS OR CHNL4);
///
///   DLDHM_CHNL5: UINT := (DLDHM OR CHNL5);
///
///   PLMDH_CHNL6: UINT := (PLMDH OR CHNL6);
///
///END_VAR
///
///PROGRAM PLC_PRG
///
///VAR
///
///END_VAR
///
///
///
///(* configure for POC *)
///
///bds_out_po_cfg(bds_out_po_signal_te.K73, STD_ACTIVE);
///
///bds_out_po_cfg(bds_out_po_signal_te.K07, STD_ACTIVE);
///
///bds_out_po_cfg(bds_out_po_signal_te.K29, STD_ACTIVE);
///
///bds_out_po_cfg(bds_out_po_signal_te.K09, STD_ACTIVE);
///
///
///
///(* configure channels for SAFOUT *)
///
///bds_safout_cfg(PHDLS_CHNL1, bds_out_po_signal_te.K73, bds_out_po_signal_te.K51, bds_out_do_signal_te.K14, 0, 0);
///
///bds_safout_cfg(DHDLM_CHNL2, bds_out_po_signal_te.K08, bds_out_do_signal_te.K16, bds_out_do_signal_te.K15, bds_out_do_signal_te.K13, 0);
///
///bds_safout_cfg(PHMDL_CHNL3, bds_out_do_signal_te.K12, bds_out_po_signal_te.K07, bds_out_po_signal_te.K29, bds_out_po_signal_te.K09, 0);
///
///bds_safout_cfg(PLDHS_CHNL4, bds_out_po_signal_te.A19, bds_out_po_signal_te.A32, bds_out_do_signal_te.A47, 0, 0);
///
///bds_safout_cfg(DLDHM_CHNL5, bds_out_po_signal_te.A03, bds_out_do_signal_te.A33, bds_out_do_signal_te.A46, bds_out_do_signal_te.A48, 0);
///
///bds_safout_cfg(PLMDH_CHNL6, bds_out_do_signal_te.A31, bds_out_po_signal_te.A05, bds_out_po_signal_te.A20, 0, 0);
///
///============================================================================
{attribute 'external_name' := 'cmp_rts_bds_safout_cfg'}
FUNCTION bds_safout_cfg : USINT
VAR_INPUT
	///The connector assigned signal name of the output.
	///
	///The channel name is composed of mode and channel number
	///
	///channel name = mode OR channel number
	///
	///and shall be defined from the application (see also example below):
	///
	///PHDLS_CHNL1: UINT := (PHDLS OR CHNL1)
	chnl_u16: UINT;
	///The common output of the channel
	outCo_u16: UINT;
	///The first output of the channel
	out1_u16: UINT;
	///The second output of the channel
	out2_u16: UINT;
	///The third output of the channel
	out3_u16: UINT;
	///The fourth output of the channel
	out4_u16: UINT;
END_VAR

END_FUNCTION

// I/O API/SAFOUT/API/bds_safout_getStatus
///Provides  status of a channel.
///
///=======
/// Remarks:
///=======
///   + The faults of the output stages are summarized in nibbels. The summarized diagnostic info looks like (see bds_safout_ts.diag_u32 and  bds_safout_ts.diag2_u32 ):
///	   + Bits   3..0		output Common
///	   + Bits   7..4		output 1
///	   + Bits   11..8		output 2
///	   + Bits 15..12		output 3
///	   + Bits 19..16		output 4
///
///   + The faults itself are defined as:
///	   + SAFOUT_SCB    	16#0001
///	   + SAFOUT_SCG    	16#0002
///	   + SAFOUT_OL     	16#0004
///	   + SAFOUT_OC     	16#0008
///
///   + Part of the status data is also the fault status of the channel DFC.
///   + With the macro function(e.g. bds_dsm_DFC_ldf) defined in DSM, the respective bit fields of the fault status can be read.
///   + bds_safout_ts.diag2_u32 provides the previous cycle(10 ms old) status of the diagnostic information. This information is not frozen and if errors are healed then it is reflected in error information. 
///
///----------
/// FFI:
///----------
///This API can be used in trusted partitions only. See Freedom from Interference (FFI) concept for more details.
///
///-----
/// Note:
///-----
///
///In mode DHDLM the current comparison between the HS and LS is not done and therefore the current deviation fault is not used. 
///
///Explanation:
///In this mode the current measurement at HS or CS at LS are not part of the functional channel (ISO25119 cat 2) but only part of the test channel.    
///
///==================================================================		  			===================================================================================================
///Return value    								  									Description
///==================================================================		  			===================================================================================================
///0																					No error.
///1																					A parameter is invalid.
///2																					Mode is wrong
///
///==================================================================		   			===================================================================================================
///
///=======
///Code Example:
///=======
///============================================================================
///
///VAR_GLOBAL CONSTANT
///
///   (* safout channel name *)
///
///   PHDLS_CHNL1: UINT := (PHDLS OR CHNL1);
///
///   DHDLM_CHNL2: UINT := (DHDLM OR CHNL2);
///
///   PHMDL_CHNL3: UINT := (PHMDL OR CHNL3);
///
///END_VAR
///
///PROGRAM PLC_PRG
///
///VAR
///
///END_VAR
///
///
///
///(* configure for POC *)
///
///bds_out_po_cfg(bds_out_po_signal_te.K73, STD_ACTIVE);
///
///bds_out_po_cfg(bds_out_po_signal_te.K07, STD_ACTIVE);
///
///bds_out_po_cfg(bds_out_po_signal_te.K29, STD_ACTIVE);
///
///bds_out_po_cfg(bds_out_po_signal_te.K09, STD_ACTIVE);
///
///
///
///(* configure channels for SAFOUT *)
///
///bds_safout_cfg(PHDLS_CHNL1, bds_out_po_signal_te.K73, bds_out_po_signal_te.K51, bds_out_do_signal_te.K14, 0, 0);
///
///bds_safout_cfg(DHDLM_CHNL2, bds_out_po_signal_te.K08, bds_out_do_signal_te.K16, bds_out_do_signal_te.K15, bds_out_do_signal_te.K13, 0);
///
///bds_safout_cfg(PHMDL_CHNL3, bds_out_do_signal_te.K12, bds_out_po_signal_te.K07, bds_out_po_signal_te.K29, bds_out_po_signal_te.K09, 0);
///
///PROGRAM appl_10ms_task
///
///VAR
///
///	chnl1_s: bds_safout_ts;
///	
///	chnl2_s: bds_safout_ts;
///	
///	chnl3_s: bds_safout_ts;
///	
///	ldf_u8: USINT := 16#00;
///
///END_VAR
///
///
///(* activate one output per channel *)
///
///bds_safout(PHDLS_CHNL1, bds_out_po_signal_te.K51, 300);
///
///bds_safout(DHDLM_CHNL2, bds_out_do_signal_te.K16, STD_ACTIVE);
///
///bds_safout(PHMDL_CHNL3, bds_out_po_signal_te.K07, 500);
///
///
///(* get status of the channels *)
///
///bds_safout_getStatus(PHDLS_CHNL1, ADR(chnl1_s));
///
///bds_safout_getStatus(DHDLM_CHNL2, ADR(chnl2_s));
///
///bds_safout_getStatus(PHMDL_CHNL3, ADR(chnl3_s));
///
///(* get last debounced fault *)
///
///ldf_u8 := bds_dsm_DFC_ldf(chnl1_s.stDFC_u16);
///
///============================================================================
{attribute 'external_name' := 'cmp_rts_bds_safout_getStatus'}
FUNCTION bds_safout_getStatus : USINT
VAR_INPUT
	///The connector assigned signal name of the output.
	///
	///The channel name is composed of mode and channel number
	///
	///channel name = mode OR channel number
	///
	///and shall be defined from the application (see also example below):
	///
	///PHDLS_CHNL1: UINT := (PHDLS OR CHNL1)
	chnl_u16: UINT;
	///Storage address of the data.
	data_ps: POINTER TO bds_safout_ts;
END_VAR

END_FUNCTION

// I/O API/SAFOUT/API/bds_safout
///Sets the output to the given state/setpoint.
///
///=======
/// Remarks:
///=======
///   + For more information also see  |bds_safout_getStatus|, |bds_safout_resetError| and |bds_safout_unlock|.
///
///----------
/// FFI:
///----------
///This API can be used in trusted partitions only. See Freedom from Interference (FFI) concept for more details.
///
///==================================================================		  			===================================================================================================
///Return value    								  									Description
///==================================================================		  			===================================================================================================
///0																					No error.
///1																					A parameter is invalid.
///2																					Mode is wrong
///3																					Output is wrong
///4																					is still locked
///5																					Requested current is out of range
///==================================================================		   			===================================================================================================
///
///=======
///Code Example:
///=======
///============================================================================
///
///VAR_GLOBAL CONSTANT
///
///   (* safout channel name *)
///
///   PHDLS_CHNL1: UINT := (PHDLS OR CHNL1);
///
///   DHDLM_CHNL2: UINT := (DHDLM OR CHNL2);
///
///   PHMDL_CHNL3: UINT := (PHMDL OR CHNL3);
///
///END_VAR
///
///PROGRAM PLC_PRG
///
///VAR
///
///END_VAR
///
///(* configure for POC *)
///
///bds_out_po_cfg(bds_out_po_signal_te.K73, STD_ACTIVE);
///
///bds_out_po_cfg(bds_out_po_signal_te.K07, STD_ACTIVE);
///
///bds_out_po_cfg(bds_out_po_signal_te.K29, STD_ACTIVE);
///
///bds_out_po_cfg(bds_out_po_signal_te.K09, STD_ACTIVE);
///
///
///(* configure channels for SAFOUT *)
///
///bds_safout_cfg(PHDLS_CHNL1, bds_out_po_signal_te.K73, bds_out_po_signal_te.K51, bds_out_do_signal_te.K14, 0, 0);
///
///bds_safout_cfg(DHDLM_CHNL2, bds_out_po_signal_te.K08, bds_out_do_signal_te.K16, bds_out_do_signal_te.K15, bds_out_do_signal_te.K13, 0);
///
///bds_safout_cfg(PHMDL_CHNL3, bds_out_do_signal_te.K12, bds_out_po_signal_te.K07, bds_out_po_signal_te.K29, bds_out_po_signal_te.K09, 0);
///
///
///PROGRAM appl_10ms_task
///
///VAR
///
///END_VAR
///
///
///(* activate one output per channel *)
///
///bds_safout(PHDLS_CHNL1, bds_out_po_signal_te.K51, 300);
///
///bds_safout(DHDLM_CHNL2, bds_out_do_signal_te.K16, STD_ACTIVE);
///
///bds_safout(PHMDL_CHNL3, bds_out_po_signal_te.K07, 500);
///
///============================================================================
{attribute 'external_name' := 'cmp_rts_bds_safout'}
FUNCTION bds_safout : USINT
VAR_INPUT
	///The connector assigned signal name of the output.
	///
	///The channel name is composed of mode and channel number
	///
	///channel name = mode OR channel number
	///
	///and shall be defined from the application (see also example below):
	///
	///PHDLS_CHNL1: UINT := (PHDLS OR CHNL1)
	chnl_u16: UINT;
	///Selected output
	out_u16: UINT;
	///State or setpoint [mA] 
	///
	///State:
	///   + STD_IDLE or STD_ACTIVE 
	///
	///Range:Based of output 
	///   + 0 to 3000 mA
	///   + 0 to 4000 mA.
	set_u16: UINT;
END_VAR

END_FUNCTION

// System API/SEC/API/bds_sec_evalRespKey
///This function is used to compare the given encrypted response key (e.g. from a diagnostic tool) with the corresponding internal stored and encrypted key for the same access level. If the keys are equal, the security manager switches to the corresponding level.
///
///=======
/// Remarks:
///=======
///   + This function can be used if the seed&key method shall be used for changing the security access level.
///   + The function |bds_sec_getSeed| must be called previously to generate a seed.
///   + This asynchronous function must be called several times until the final result is available.
///   + This function will be rejected if another asynchronous security function was already started for this instance.
///   + After a reset, this function can be executed successfully after 500ms at the earliest.
///   + The completion of this function (execution within a loop) takes about 90us (microseconds) if there is no HSM access conflict with another instance.
///   + For each retry of this function a new seed must be requested with function |bds_sec_getSeed|.  
///
///----------
/// FFI:
///----------
///This API can be used in trusted partitions only. See Freedom from Interference (FFI) concept for more details.
///
///-----
/// Info:
///-----
///
///If the function has been called 3 times with an incorrect key, the function is locked for security reasons until the next ECU reset.
///
///==================================================================		  			===================================================================================================
///Return value    								  									Description
///==================================================================		  			===================================================================================================
///16#0000: BDS_SEC_ERR_NO_ERROR_DU16													Function was executed without errors. The requested security access level is unlocked.
///16#0001: BDS_SEC_ERR_PARAM1_ERROR_DU16												Invalid instance number
///16#0002: BDS_SEC_ERR_PARAM2_ERROR_DU16												Invalid access level
///16#0003: BDS_SEC_ERR_PARAM3_ERROR_DU16												Invalid response key pointer. Pointer is equal to zero
///16#0010: BDS_SEC_ERR_REQUEST_PENDING_DU16											This asynchronous function was not yet completed and must be called again with the same parameter values. Several function calls may be required in particular if another security manager instance is also running
///16#0011: BDS_SEC_ERR_WAIT_FOR_STARTUP_DELAY_DU16										The mandatory start up delay of 500ms has not yet expired. Repeat the function call after some time
///16#0020: BDS_SEC_ERR_INVALID_SEQUENCE_DU16											This function was called without requesting a seed previously with bds_sec_getSeed or although another asynchronous security function was not yet completed. The other asynchronous function that has already been started must be called again and must be completed before this function can be started
///16#0021: BDS_SEC_ERR_NBR_ATTEMPTS_EXCEEDED_DU16										The maximum number of function calls with an incorrect response key has been reached. A restart is required for further attempts
///16#0033: BDS_SEC_ERR_OPEN_SESSION_FAILED_DU16										Security session could not be opened for this functionPossible reason could be that the HSM is not running
///16#0034: BDS_SEC_ERR_GENERATE_RANDOM_FAILED_DU16										The process to generate the random has been failed
///16#0035: BDS_SEC_ERR_CLOSE_SESSION_FAILED_DU16										Security session could not be closed for this function
///16#0036: BDS_SEC_ERR_ENCRYPT_INIT_FAILED_DU16										Internal encryption initialization has been failed. To terminate the function, it must be called again
///16#0037: BDS_SEC_ERR_ENCRYPT_FAILED_DU16												Internal encrypt operation has been failed. To terminate the function, it must be called again
///16#0039: BDS_SEC_ERR_COMPARE_KEY_FAILED_DU16											The given response key does not match with the internal calculated key or the execution of the function was aborted due to an error. The current access level remains unchanged
///
///==================================================================		   			===================================================================================================
///
///For Access levels, Refer the below table & provide the value,
///
///==================================================================		  			===================================================================================================
///Access Level Variable   								  							Value
///==================================================================		  			===================================================================================================
///BDS_SEC_ACC_LEVEL_0_E																0
///BDS_SEC_ACC_LEVEL_1_E																1
///BDS_SEC_ACC_LEVEL_2_E																2
///BDS_SEC_ACC_LEVEL_3_E																3
///BDS_SEC_ACC_LEVEL_4_E																4
///BDS_SEC_ACC_LEVEL_5_E																5
///BDS_SEC_ACC_LEVEL_6_E																6
///BDS_SEC_ACC_LEVEL_7_E																7
///BDS_SEC_ACC_LEVEL_8_E																8
///BDS_SEC_ACC_LEVEL_9_E																9
///BDS_SEC_ACC_LEVEL_10_E																10
///BDS_SEC_ACC_LEVEL_11_E																11
///BDS_SEC_ACC_LEVEL_12_E																12
///BDS_SEC_ACC_LEVEL_13_E																13
///BDS_SEC_ACC_LEVEL_14_E																14
///BDS_SEC_ACC_LEVEL_15_E																15
///BDS_SEC_ACC_LEVEL_16_E																16
///BDS_SEC_ACC_LEVEL_17_E																17
///BDS_SEC_ACC_LEVEL_18_E																18
///BDS_SEC_ACC_LEVEL_19_E																19
///BDS_SEC_ACC_LEVEL_20_E																20
///
///==================================================================		   			===================================================================================================
///=======
///Code Example:
///=======
///============================================================================
///
///PROGRAM appl_Task_1
///
///  VAR
///	return_u16 : UINT;
///
///	respKey_au8 : ARRAY[0..15] OF USINT;
///	
///  END_VAR
///  
///  (*evaluate the response key*)
///  
///result_u16 := bds_sec_evalRespKey(bds_diag_inst_te.BDS_SEC_ASW_INST_NAME_1_E, 2, ADR(respKey_au8));
///  
///============================================================================
{attribute 'external_name' := 'cmp_rts_bds_sec_evalRespKey'}
FUNCTION bds_sec_evalRespKey : UINT
VAR_INPUT
	///Instance number. pointer to |bds_diag_inst_te|
	diagInst_e: bds_diag_inst_te;
	///The new access level. Refer access level table
	level_e: USINT;
	///Pointer to a 16 byte buffer must be declared in the application and must contain the response key from diagnostic tool for comparision.
	respKey_pau8: POINTER TO USINT;
END_VAR

END_FUNCTION

// System API/SEC/API/bds_sec_getSeed
///This function is used to request a seed value (random Number with 128Bit). The random number is generated by the Hardware Security Module (HSM) of the RC.
///
///=======
/// Remarks:
///=======
///
///   + This function can be used if the seed&key method shall be used for changing the security access level.
///   + After successful execution of this function the generated seed will be also internally stored for a following key compare with |bds_sec_evalRespKey|.
///   + This asynchronous function must be called several times until the final result is available.
///   + The completion of this function (execution within a loop) takes about 50us (microseconds) if there is no HSM access conflict with another instance.
///   + This function will be rejected if another asynchronous security function was already started for this instance.
///
///----------
/// FFI:
///----------
///This API can be used in trusted partitions only. See Freedom from Interference (FFI) concept for more details.
///
///==================================================================		  			===================================================================================================
///Return value    								  									Description
///==================================================================		  			===================================================================================================
///16#0000:BDS_SEC_ERR_NO_ERROR_DU16													Function was executed without errors. The requested seed was copied to the given buffer.
///16#0001: BDS_SEC_ERR_PARAM1_ERROR_DU16												Invalid instance number. 
///16#0002: BDS_SEC_ERR_PARAM2_ERROR_DU16												Invalid seed pointer. Pointer is equal to zero.
///16#0010: BDS_SEC_ERR_REQUEST_PENDING_DU16											This asynchronous function was not yet completed and must be called again with the same parameter values. Several function calls may be required in particular if another security manager instance is also running.
///16#0020:BDS_SEC_ERR_INVALID_SEQUENCE_DU16											This function was called although another asynchronous security function was not yet completed. The other asynchronous function that has already been started must be called again and must be completed before this function can be started.
///16#0033: BDS_SEC_ERR_OPEN_SESSION_FAILED_DU16										Security session could not be opened for this function. Possible reason could be that the HSM is not running.
///16#0034: BDS_SEC_ERR_GENERATE_RANDOM_FAILED_DU16									The process to generate the random has been failed. To terminate the function, it must be called again.
///16#0035: BDS_SEC_ERR_CLOSE_SESSION_FAILED_DU16										Security session could not be closed for this function. 
///
///==================================================================		   			===================================================================================================
///=======
///Code Example:
///=======
///============================================================================
///
///PROGRAM appl_Task_1
///
///  VAR
///	return_u16 : UINT;
///
///	seed_au8 : ARRAY[0..15] OF USINT;
///	
///  END_VAR
///
///return_u16 := bds_sec_getSeed(bds_diag_inst_te.BDS_SEC_ASW_INST_NAME_1_E, ADR(seed_au8));
///  
///============================================================================
///
{attribute 'external_name' := 'cmp_rts_bds_sec_getSeed'}
FUNCTION bds_sec_getSeed : UINT
VAR_INPUT
	///Instance number . pointer to |bds_diag_inst_te|
	diagInst_e: bds_diag_inst_te;
	///Pointer to a 16 byte buffer which must be provided by the application. Generated seed will be copied to this buffer.
	seed_pau8: POINTER TO USINT;
END_VAR

END_FUNCTION

// System API/SEC/API/bds_sec_getLevel
///This API function is used to get the current security access level for a specific security instance.
///
///=======
/// Remarks:
///=======
///
///   + This function reads the security level which was previously set with functions |bds_sec_setLevel| or |bds_sec_evalRespKey|.
///
///----------
/// FFI:
///----------
///This API can be used in trusted partitions only. See Freedom from Interference (FFI) concept for more details.
///
///==================================================================		  			===================================================================================================
///Return value    								  									Description
///==================================================================		  			===================================================================================================
///16#0000: BDS_SEC_ERR_NO_ERROR_DU16													Function was executed without errors
///16#0001:  BDS_SEC_ERR_PARAM1_ERROR_DU16												Invalid instance number. 
///16#0002: BDS_SEC_ERR_PARAM2_ERROR_DU16												Invalid access level pointer. Pointer is equal to zero
///
///==================================================================		   			===================================================================================================
///
///For Access levels, Refer the below table & provide the value,
///
///==================================================================		  			===================================================================================================
///Access Level Variable   								  							Value
///==================================================================		  			===================================================================================================
///BDS_SEC_ACC_LEVEL_0_E																0
///BDS_SEC_ACC_LEVEL_1_E																1
///BDS_SEC_ACC_LEVEL_2_E																2
///BDS_SEC_ACC_LEVEL_3_E																3
///BDS_SEC_ACC_LEVEL_4_E																4
///BDS_SEC_ACC_LEVEL_5_E																5
///BDS_SEC_ACC_LEVEL_6_E																6
///BDS_SEC_ACC_LEVEL_7_E																7
///BDS_SEC_ACC_LEVEL_8_E																8
///BDS_SEC_ACC_LEVEL_9_E																9
///BDS_SEC_ACC_LEVEL_10_E																10
///BDS_SEC_ACC_LEVEL_11_E																11
///BDS_SEC_ACC_LEVEL_12_E																12
///BDS_SEC_ACC_LEVEL_13_E																13
///BDS_SEC_ACC_LEVEL_14_E																14
///BDS_SEC_ACC_LEVEL_15_E																15
///BDS_SEC_ACC_LEVEL_16_E																16
///BDS_SEC_ACC_LEVEL_17_E																17
///BDS_SEC_ACC_LEVEL_18_E																18
///BDS_SEC_ACC_LEVEL_19_E																19
///BDS_SEC_ACC_LEVEL_20_E																20
///
///==================================================================		   			===================================================================================================
///=======
///Code Example:
///=======
///============================================================================
///
///PROGRAM appl_Task_1
///
///  VAR
///	return_u16 : UINT;
///
///	secLevel: POINTER TO USINT;
///
///  END_VAR
///
///(*get the actual access level*)
///
///return_u16 := bds_sec_getLevel(bds_diag_inst_te.BDS_SEC_ASW_INST_NAME_1_E, ADR(secLevel));
///  
///============================================================================
{attribute 'external_name' := 'cmp_rts_bds_sec_getLevel'}
FUNCTION bds_sec_getLevel : UINT
VAR_INPUT
	///Instance number. pointer to |bds_diag_inst_te|
	diagInst_e: bds_diag_inst_te;
	///Pointer to a variable which must be provided(Refer access level table). The current level will be copied to this variable. 
	actLevel_pe: POINTER TO USINT;
END_VAR

END_FUNCTION

// System API/SEC/API/bds_sec_setLevel
/// This API function is used to set the security access level.
///
///=======
/// Remarks:
///=======
///
///   + This function sets the security access level directly without any seed&key procedure. 
///   + The function can be used if the security access is directly controlled by the application
///
///----------
/// FFI:
///----------
///This API can be used in trusted partitions only. See Freedom from Interference (FFI) concept for more details.
///
///==================================================================		  			===================================================================================================
///Return value    								  									Description
///==================================================================		  			===================================================================================================
///16#0000: BDS_SEC_ERR_NO_ERROR_DU16													Function was executed without errors
///16#0001: BDS_SEC_ERR_PARAM1_ERROR_DU16												Invalid instance number
///16#0002: BDS_SEC_ERR_PARAM2_ERROR_DU16												Invalid access level
///
///==================================================================		   			===================================================================================================
///
///For Access levels, Refer the below table & provide the value,
///
///==================================================================		  			===================================================================================================
///Access Level Variable   								  							Value
///==================================================================		  			===================================================================================================
///BDS_SEC_ACC_LEVEL_0_E																0
///BDS_SEC_ACC_LEVEL_1_E																1
///BDS_SEC_ACC_LEVEL_2_E																2
///BDS_SEC_ACC_LEVEL_3_E																3
///BDS_SEC_ACC_LEVEL_4_E																4
///BDS_SEC_ACC_LEVEL_5_E																5
///BDS_SEC_ACC_LEVEL_6_E																6
///BDS_SEC_ACC_LEVEL_7_E																7
///BDS_SEC_ACC_LEVEL_8_E																8
///BDS_SEC_ACC_LEVEL_9_E																9
///BDS_SEC_ACC_LEVEL_10_E																10
///BDS_SEC_ACC_LEVEL_11_E																11
///BDS_SEC_ACC_LEVEL_12_E																12
///BDS_SEC_ACC_LEVEL_13_E																13
///BDS_SEC_ACC_LEVEL_14_E																14
///BDS_SEC_ACC_LEVEL_15_E																15
///BDS_SEC_ACC_LEVEL_16_E																16
///BDS_SEC_ACC_LEVEL_17_E																17
///BDS_SEC_ACC_LEVEL_18_E																18
///BDS_SEC_ACC_LEVEL_19_E																19
///BDS_SEC_ACC_LEVEL_20_E																20
///
///==================================================================		   			===================================================================================================
///
///=======
///Code Example:
///=======
///============================================================================
///
///PROGRAM appl_Task_1
///
///  VAR
///
///	return_u16 : UINT;
///
///  END_VAR
///
///  (*set a new access level*)
///  
///return_u16 := bds_sec_setLevel(bds_diag_inst_te.BDS_SEC_ASW_INST_NAME_1_E, 2);
///  
///============================================================================
///
{attribute 'external_name' := 'cmp_rts_bds_sec_setLevel'}
FUNCTION bds_sec_setLevel : UINT
VAR_INPUT
	///Instance number. pointer to |bds_diag_inst_te|
	diagInst_e: bds_diag_inst_te;
	///Pointer to a variable which must be provided(Refer access level table). The current level will be copied to this variable. 
	newLevel_e: USINT;
END_VAR

END_FUNCTION

// System API/SEC/API/bds_sec_getRnd
///This API function is used to generate a random number. The random number is generated by the Hardware Security Module (HSM) of the RC.
///
///=======
/// Remarks:
///=======
///
///   + This random number can be freely used by the application. It is independent of the implemented seed&key method.
///   + This asynchronous function must be called several times until the final result is available.
///   + At least one function call is required per 16 bytes of the random number.
///   + Each generation of 16 bytes of the random number takes about 40us (microseconds) if there is no HSM access conflict with another instance.
///   + This function will be rejected if it was already started but not yet finished with another buffer pointer.
///
///----------
/// FFI:
///----------
///This API can be used in trusted partitions only. See Freedom from Interference (FFI) concept for more details.
///
///==================================================================		  			===================================================================================================
///Return value    								  									Description
///==================================================================		  			===================================================================================================
///16#0000:BDS_SEC_ERR_NO_ERROR_DU16													Function was executed without errors
///16#0001: BDS_SEC_ERR_PARAM1_ERROR_DU16												Invalid buffer pointer. Pointer is equal to zero.
///16#0002: BDS_SEC_ERR_PARAM2_ERROR_DU16												Invalid size. See parameter description.
///16#0010: BDS_SEC_ERR_REQUEST_PENDING_DU16											This asynchronous function was not yet completed and must be called again with the same parameter values. Several function calls may be required in particular if another security manager instance is also running.
///16#0020:BDS_SEC_ERR_INVALID_SEQUENCE_DU16											This function was called with another buffer pointer although the function with the previous buffer pointer was not yet completed. The function has to be called again with the previous buffer pointer until completion before it can be started with a new buffer pointer.
///16#0033: BDS_SEC_ERR_OPEN_SESSION_FAILED_DU16										Security session could not be opened for this function.Possible reason could be that the HSM is not running. 
///16#0034: BDS_SEC_ERR_GENERATE_RANDOM_FAILED_DU16										The process to generate the random has been failed. To terminate the function, it must be called again.
///16#0035: BDS_SEC_ERR_CLOSE_SESSION_FAILED_DU16										Security session could not be closed for this function. 
///
///==================================================================		   			===================================================================================================
///
///=======
///Code Example:
///=======
///============================================================================
///
///PROGRAM appl_Task_1
///
///  VAR
///
///	return_u16 : UINT;
///
///	RND_SIZE_DU16 : UINT := 100;
///
///	rnd_au8 : ARRAY[0..99] OF USINT;
///
///  END_VAR
///
///(*check for request to generate a new random*)
///
///return_u16 := bds_sec_getRnd(ADR(rnd_au8), RND_SIZE_DU16);
///  
///============================================================================
///
{attribute 'external_name' := 'cmp_rts_bds_sec_getRnd'}
FUNCTION bds_sec_getRnd : UINT
VAR_INPUT
	///Pointer to a buffer (buffer size = size_u16) which must be provided by the application. Generated random number will be copied to this buffer.
	buf_pau8: POINTER TO USINT;
	///Size [in bytes] of the requested random number and of the buffer above.
	///
	///Value range:1..512
	size_u16: UINT;
END_VAR

END_FUNCTION

// System API/SEC/API/bds_sec_resetLevel
/// This API function is used to reset the security access level to the DEFAULT level.
///
///=======
/// Remarks:
///=======
///
///This functions resets the security level which was previously set with functions |bds_sec_setLevel| or |bds_sec_evalRespKey|.
///
///----------
/// FFI:
///----------
///This API can be used in trusted partitions only. See Freedom from Interference (FFI) concept for more details.
///
///==================================================================		  			===================================================================================================
///Return value    								  									Description
///==================================================================		  			===================================================================================================
///16#0000: BDS_SEC_ERR_NO_ERROR_DU16													Function was executed without errors
///16#0001: BDS_SEC_ERR_PARAM1_ERROR_DU16												Invalid instance number. 
///
///==================================================================		   			===================================================================================================
///=======
///Code Example:
///=======
///============================================================================
///
///PROGRAM appl_Task_1
///
///  VAR
///
///	return_u16 : UINT;
///
///  END_VAR
///
///  (*reset to default level*)
///  
///return_u16 := bds_sec_resetLevel(bds_diag_inst_te.BDS_SEC_ASW_INST_NAME_1_E);
///
///============================================================================
///
{attribute 'external_name' := 'cmp_rts_bds_sec_resetLevel'}
FUNCTION bds_sec_resetLevel : UINT
VAR_INPUT
	///Instance number. pointer to |bds_diag_inst_te|
	diagInst_e: bds_diag_inst_te;
END_VAR

END_FUNCTION

